Staubli VAL3: CurrentTool.pjx

--- CurrentTool.pjx ---
Parameters version=s8.8.3Cs9_BS1660 stackSize=5000 millimeterUnit=true
Data file=CurrentTool.dtx

--- CurrentTool.dtx ---
public num nItem
public tool tValue = {fatherId=flange[0]}
public string sName
public num nItemM
